(* PLC project Line.project, CODESYS CODESYS V3.5 SP19 *)
(* stored: creationDateTime 2026-10-19T10:00:00, modificationDateTime 2026-10-19T10:00:00 *)

VAR_GLOBAL  (* GVL_IO *)
  xLampOut AT %QX0.0 : BOOL;
END_VAR

{attribute 'hide_all_locals'}
FUNCTION_BLOCK FB_Average EXTENDS FB_Base IMPLEMENTS I_Value
VAR_INPUT
	nSize : INT := 10; // window
END_VAR
VAR
	aValues : ARRAY[1..10] OF REAL;
	nCount : INT;
END_VAR

            IF nCount < nSize THEN
	nCount := nCount + 1;
END_IF
          

METHOD Add : BOOL
  VAR_INPUT
    rValue : REAL;
  END_VAR
                  aValues[nCount] := rValue;
Add := TRUE;
                
END_METHOD

PROPERTY Count : INT
GET
Count := nCount;
END_GET
END_PROPERTY
END_FUNCTION_BLOCK

{attribute 'qualified_only'}
PROGRAM PLC_PRG
  VAR
    xStart : BOOL;
    xStop : BOOL;
    xMotor : BOOL;
    fbBlink : BLINK;
    rIn : REAL;
    rOut : REAL;
  END_VAR
  VAR  (* added by the conversion: wires and edge detectors of the diagram *)
    _w4 : BOOL;
    _w5 : BOOL;
  END_VAR

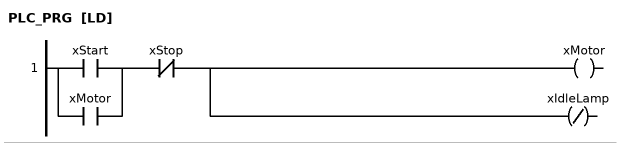
(* LD diagram, written out as Structured Text *)

_w4 := xMotor;
_w5 := (xStart OR _w4) AND NOT xStop;
xMotor := _w5;
xIdleLamp := NOT _w5;

ACTION Scale:
(* FBD diagram, written out as Structured Text *)
rOut := rIn * 2.5;
fbBlink(EN := xMotor, ENABLE := xMotor);
END_ACTION
END_PROGRAM

CONFIGURATION Device
  RESOURCE Application ON PLC
    TASK MainTask(PRIORITY := 1);
    PROGRAM PLC_PRG WITH MainTask : PLC_PRG;
  END_RESOURCE
END_CONFIGURATION
